Fanuc KAREL source: ka00155.KL

PROGRAM KA00155
%STACKSIZE=65535
%PRIORITY=65535
%NOLOCKGROUP
VAR
SRC : ARRAY[4] OF REAL
DST : ARRAY[4] OF REAL
BEGIN
-- UNRESOLVED_PC line 7 opcodes [22 22 1E] marker_code=0
END KA00155
